(* IEC 61131-3 sources: llm-plc-st-eval/data/processed_definitivo/gpt-4o-2024-08-06/I6/few_shot, 3 files *)

(* ---- ejec_1.st ---- *)
FUNCTION_BLOCK FB_Temperatura
VAR_INPUT
    rawTemp : INT; (* Señal de temperatura cruda *)
END_VAR
VAR_OUTPUT
    tempC : REAL; (* Temperatura en grados Celsius *)
    enfriador : BOOL; (* Estado del enfriador *)
    almSensor : BOOL; (* Alarma de sensor *)
END_VAR
VAR
    tempC_prev : REAL; (* Valor previo de tempC para histéresis *)
END_VAR

(* Convertir rawTemp a grados Celsius *)
tempC := (REAL(rawTemp) * 100.0) / 27648.0;

(* Comprobar si rawTemp está fuera de rango *)
IF (rawTemp < 0) OR (rawTemp > 27648) THEN
    almSensor := TRUE;
    enfriador := FALSE;
ELSE
    almSensor := FALSE;

    (* Control del enfriador con histéresis *)
    IF tempC >= 80.0 THEN
        enfriador := TRUE;
    ELSIF tempC <= 75.0 THEN
        enfriador := FALSE;
    ELSE
        enfriador := enfriador; (* Mantener el estado actual *)
    END_IF;
END_IF;

END_FUNCTION_BLOCK

(* ---- ejec_2.st ---- *)
FUNCTION_BLOCK FB_Temperatura
VAR_INPUT
    rawTemp : INT; (* Señal de temperatura cruda *)
END_VAR
VAR_OUTPUT
    tempC : REAL; (* Temperatura en grados Celsius *)
    enfriador : BOOL; (* Estado del enfriador *)
    almSensor : BOOL; (* Alarma del sensor *)
END_VAR
VAR
    tempC_prev : REAL; (* Temperatura previa para histéresis *)
END_VAR

(* Verificar si la señal de temperatura está fuera de rango *)
IF (rawTemp < 0) OR (rawTemp > 27648) THEN
    almSensor := TRUE;
    enfriador := FALSE;
ELSE
    almSensor := FALSE;

    (* Calcular la temperatura en grados Celsius *)
    tempC := (REAL(rawTemp) * 100.0) / 27648.0;

    (* Control del enfriador con histéresis *)
    IF tempC >= 80.0 THEN
        enfriador := TRUE;
    ELSIF tempC <= 75.0 THEN
        enfriador := FALSE;
    ELSE
        enfriador := enfriador; (* Mantener el estado actual *)
    END_IF;
END_IF;
END_FUNCTION_BLOCK

(* ---- ejec_3.st ---- *)
FUNCTION_BLOCK FB_Temperatura
VAR_INPUT
    rawTemp : INT; (* Señal de temperatura cruda *)
END_VAR
VAR_OUTPUT
    tempC : REAL; (* Temperatura en grados Celsius *)
    enfriador : BOOL; (* Estado del enfriador *)
    almSensor : BOOL; (* Alarma del sensor *)
END_VAR
VAR
    tempC_prev : REAL; (* Valor previo de tempC para histéresis *)
END_VAR

(* Convertir rawTemp a grados Celsius *)
tempC := (REAL(rawTemp) * 100.0) / 27648.0;

(* Verificar si rawTemp está fuera de rango *)
IF (rawTemp < 0) OR (rawTemp > 27648) THEN
    almSensor := TRUE;
    enfriador := FALSE;
ELSE
    almSensor := FALSE;

    (* Control del enfriador con histéresis *)
    IF tempC >= 80.0 THEN
        enfriador := TRUE;
    ELSIF tempC <= 75.0 THEN
        enfriador := FALSE;
    ELSE
        enfriador := enfriador; (* Mantener estado actual *)
    END_IF;
END_IF;

END_FUNCTION_BLOCK
